// TIA Portal V21 export
// export: Created 2026-11-18T04:30:50.1315089Z, ExportSetting WithDefaults, DisplayName Totally Integrated Automation Portal, DisplayVersion V21, DisplayName STEP 7 Professional, DisplayVersion V21, DisplayName STEP 7 Safety, DisplayVersion V21, DisplayName Tech WebApplication, DisplayVersion V21, DisplayName WinCC Basic/Comfort/Advanced, DisplayVersion V21
TagTable "Tags_Line_Control"
  HMI_Btn_Start : Bool  (1 s)
  HMI_Btn_Stop : Bool  (1 s)
  HMI_Btn_Reset_Alarm : Bool  (1 s)
  HMI_Btn_Reset_Counter : Bool  (1 s)
  HMI_Sw_Mode_Auto : Bool  (1 s)
  PLC_Sys_Status : Int  (1 s)
  PLC_Conveyor_Run : Bool  (1 s)
  PLC_VJ_Printer_Ready : Bool  (1 s)
  PLC_Cognex_Sensor_Trig : Bool  (1 s)
  PLC_Cognex_Sensor_Count : DInt  (1 s)
  PLC_Cognex_Status : Int  (1 s)
  PLC_Label_Sensor_Trig : Bool  (1 s)
  PLC_Label_Sensor_Count : DInt  (1 s)
  PLC_Labeller_Active : Bool  (1 s)
  PLC_Keyence_Status : Int  (1 s)
  PLC_Reject_Sensor_Trig : Bool  (1 s)
  PLC_Reject_Sensor_Count : DInt  (1 s)
  PLC_Rejecter_Actuated : Bool  (1 s)
  PLC_Total_Reject_Count : DInt  (1 s)
  PLC_Scanner_Status_1 : Int  (1 s)
  PLC_Scanner_Status_2 : Int  (1 s)
  PLC_Scanner_Status_3 : Int  (1 s)
  PLC_Alm_Missing_Prod : Bool  (1 s)
  PLC_ID_Status_1 : Int  (1 s)
  PLC_ID_Status_2 : Int  (1 s)
  PLC_ID_Status_3 : Int  (1 s)
  PLC_ID_Status_4 : Int  (1 s)
  PLC_ID_Status_5 : Int  (1 s)
  PLC_ID_Status_6 : Int  (1 s)
  PLC_ID_Status_7 : Int  (1 s)
  PLC_ID_Status_8 : Int  (1 s)
